FUNCTION WRITE_PROTECTED_INT
VAR_INPUT
    Ptr : POINTER TO INT;
    Value : INT;
END_VAR

Ptr^ := Value;

END_FUNCTION

(* stored: Version 1.1.0.1
   POU WRITE_PROTECTED_INT: Id {d5d23a20-8f67-4a43-b9e4-bf7852dc7164}, SpecialFunc None *)
